Fanuc KAREL source: ko00071.KL

PROGRAM KO00071
%STACKSIZE=65535
%PRIORITY=65535
%NOLOCKGROUP
VAR
P1 : XYZWPREXT
P2 : XYZWPR
F : BOOLEAN
OUT : XYZWPREXT
BEGIN
F=TRUE
-- UNSAFE_SOURCE_IR line 11: OUT = MIRROR(P1, convert_xyzwpr_to_position(P2), F)
END KO00071
